Fanuc KAREL source: kb00033.KL

-- PROVISIONAL review KL for V770-1; original PC SHA256 bc2e66a77dc4f2291affe1675c8a3a49c4e0c2b70e0973a9e12f2954d5e582ee
-- Incomplete behavior may be omitted. Consult companion uncertainty JSON. Do not deploy.
PROGRAM KB00033
%NOLOCKGROUP
BEGIN
  -- UNRESOLVED_PC offsets 5-14; opcodes 3F,75
  -- UNRESOLVED_PC offsets 19-26; opcodes 9D,23
  -- UNRESOLVED_PC offsets 31-57; opcodes 27,22,22,2A,22,27,9D,31
  -- UNRESOLVED_PC offsets 62-66; opcodes 7F
END KB00033
